Fanuc KAREL source: kd00036.KL

-- PROVISIONAL review KL for V1013-1; original PC SHA256 872a5c9b6268101cc24685c1f9c048bbf0eee64f8f7980d60d47e5499ca85833
-- Incomplete behavior may be omitted. Consult companion uncertainty JSON. Do not deploy.
PROGRAM KD00036
%NOLOCKGROUP
VAR
  I : INTEGER
  J : INTEGER
  B : BOOLEAN
  R : REAL
  S : STRING[80]
BEGIN
  -- UNRESOLVED_PC offsets 5-17; opcodes 9D,81,18,9D,1B,9D,12,13,04
  -- UNRESOLVED_PC offsets 22-26; opcodes 7F
END KD00036
